RoboDK station: Robot_2_2025.rdk

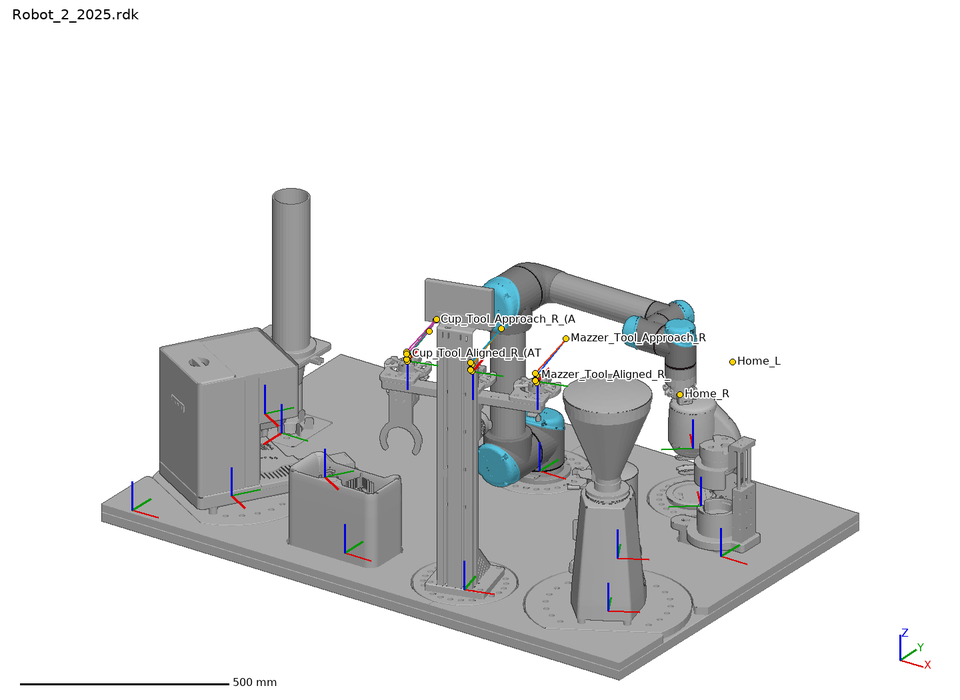
[picture v0: the station drawn from its stored meshes, robots at their saved joint values, targets as dots, program paths as lines]
Station Robot_2_2025 (saved by RoboDK 6.0.7). Poses are relative to the parent item; angles as X-Y-Z fixed-axis rotations.
Station parameters (name, value as stored): IO_5, 1, IO_2, 0, IO_3, 0, IO_4, 0, IO_1, 0, IO_0, 0, 0, 0, 1, 0, 4, 0
  - frame UR5_Base at (0, 0, 0) mm
    - robot UR5: 6 axes
        modified DH rows (alpha deg, a mm, theta deg, d mm): 0, 0, 0, 89.2; 90, 0, 180, 0; 0, 425, 0, 0; 0, 392, 0, 109.3; -90, 0, 0, 94.75; 90, 0, 180, 82.5
        joint limits [-360, -360, -360, -360, -360, -360] to [360, 360, 360, 360, 360, 360]; home [0, -90, -90, 0, 90, 0]; saved at [-0.001, -89.995, -89.998, -90.003, 89.998, 0.001]
      - tool Master_Tool_(UR5), TCP at (0, 0, 48.94) mm, size 88.9 x 94.7 x 67.9 mm
      - tool Cup_Tool_Shut_(UR5), TCP at (-34.39, 40.98, 235.56) mm, rotated rx 0 ry 0 rz -50 deg, size 116 x 104.2 x 218.8 mm
      - tool Cup_Tool_Open_(UR5), TCP at (-67.17, 80.05, 235.56) mm, rotated rx 0 ry 0 rz -50 deg, size 166.5 x 104.2 x 218.8 mm
      - tool Mazzer_Tool_(UR5), TCP at (0, 0, 153.18) mm, rotated rx 0 ry 0 rz -50 deg, size 105.5 x 104.2 x 106.6 mm
      - tool Rancilio_Tool_(UR5), TCP at (18.19, -21.68, 194.84) mm, rotated rx 0 ry -3.9 rz -50 deg, size 87.5 x 104.2 x 184.8 mm
      - tool Cup_(UR5), TCP at (-82.31, 98.09, 235.54) mm, rotated rx 0 ry 0 rz -50 deg, size 79 x 78 x 79 mm
    - object UR5_Plate at (0, 0, 0) mm, size 249.9 x 249.9 x 20 mm, geometry from UR5_Plate.STL
    - frame Table_Top at (-700, -700, -20) mm
      - object Table_Top at (0, 0, 0) mm, size 1515 x 1000 x 25 mm, geometry from Table_Top.STL
      - object Table_Cushion at (0, 0, 0) mm, size 1515 x 1000 x 20 mm, geometry from Table_Cushion.STL
      - frame Rancilio at (150, 200, 0) mm, rotated rx 0 ry 0 rz -30 deg
        - object Rancilio at (0, 0, 0) mm, size 399.6 x 458 x 388.3 mm, geometry from Rancilio_Assembly.STL
        - frame Rancilio_Tool at (39.29, 69.7, 222) mm
          - object Rancilio_Tool_Inserted_(Rancilio) at (0, 0, 0) mm, rotated rx 0 ry -90 rz 45 deg, size 87.1 x 104.3 x 184.1 mm, geometry from Rancilio_Tool_Assembly.STL
          - object Rancilio_Tool_Rotated_(Rancilio) at (0, 0, 0) mm, rotated rx 0 ry -90 rz 75 deg, size 87.1 x 104.3 x 184.1 mm, geometry from Rancilio_Tool_Assembly.STL
        - frame Rancilio_Scale at (39, 226.92, 20) mm
          - object Cup_(Rancilio) at (0, -157.52, 65.24) mm, size 79 x 79 x 78 mm, geometry from Supreme_Cup.STL
          - object Rancilio_Scale_Lock at (0, 0, 0) mm, size 100.1 x 260 x 71.4 mm, geometry from Rancilio_Scale_Assembly_1_Lock.STL
          - object Rancilio_Scale_Read at (0, 0, 0) mm, size 100.1 x 260 x 71.4 mm, geometry from Rancilio_Scale_Assembly_1_Read.STL
      - frame Rancilio_Tool_Cleaner at (550, 100, 0) mm
        - object Rancilio_Tool_Cleaner at (0, 0, 0) mm, size 258 x 136.9 x 218.7 mm, geometry from Portafilter_Cleaner_Assembly.STL
      - frame ATI at (900, 100, 0) mm, rotated rx 0 ry 0 rz 15 deg
        - object ATI at (0, 0, 0) mm, size 444.3 x 250 x 843.3 mm, geometry from ATI_Assembly_1.STL
        - frame Cup_Tool_(ATI) at (-163.9, 54.25, 556) mm, rotated rx 180 ry 0 rz 90 deg
          - object Cup_Tool_Shut_(ATI) at (0, 0, 0) mm, size 116 x 104.3 x 218.9 mm, geometry from Cup_Tool_Assembly_Closed.STL
          - target Cup_Tool_Approach_R_(ATI) (joint target) at (200, -1, -18) mm, rotated rx 0 ry 0 rz 50 deg; joints [-77.671, -81.541, -71.804, -116.654, 90.001, -222.671] of UR5
          - target Cup_Tool_Aligned_R_(ATI) (joint target) at (0.64, -1.17, -18.29) mm, rotated rx -0.48 ry 0.34 rz 50.01 deg; joints [-76.902, -110.177, -39.589, -120.099, 90.575, -221.892] of UR5
          - target Cup_Tool_Inserted_R_(ATI) (joint target) at (1.17, -1.09, 0) mm, rotated rx -0.52 ry 0.38 rz 50.08 deg; joints [-76.908, -108.351, -45.194, -116.323, 90.631, -221.828] of UR5
          - target Cup_Tool_Mated_R_(ATI) (joint target) at (0.72, -1.18, 0.85) mm, rotated rx -0.51 ry 0.38 rz 50.07 deg; joints [-76.914, -108.36, -45.32, -116.191, 90.623, -221.837] of UR5
          - target Cup_Tool_Attached_R_(ATI) (joint target) at (1.05, -1.02, -11) mm, rotated rx -0.5 ry 0.36 rz 50.03 deg; joints [-76.894, -109.363, -41.97, -118.536, 90.601, -221.86] of UR5
          - target Cup_Tool_Rotated_R_(ATI) (joint target) at (1.07, -1.03, -11.05) mm, rotated rx 0.35 ry 0.5 rz 140.04 deg; joints [-76.895, -109.361, -41.967, -118.536, 90.599, -131.856] of UR5
          - target Cup_Tool_Departure_R_(ATI) (joint target) at (151, -1, -11) mm, rotated rx 0 ry 0 rz 140 deg; joints [-77.368, -87.366, -67.792, -114.84, 90.001, -132.368] of UR5
          - target Cup_Tool_Approach_L_(ATI) (joint target) at (200, 0, -20) mm, rotated rx 0 ry 0 rz 50.44 deg; joints [70.564, -98.372, 71.405, -63.033, -89.998, -254] of UR5
          - target Cup_Tool_Aligned_L_(ATI) (joint target) at (2.26, -4.72, -23.42) mm, rotated rx -0.9 ry 0.14 rz 50.33 deg; joints [81.304, -69.621, 38.471, -59.135, -89.129, -243.367] of UR5
          - target Cup_Tool_Inserted_L_(ATI) (joint target) at (2, -4.79, -4.65) mm, rotated rx -0.97 ry 0.67 rz 50.05 deg; joints [81.242, -71.217, 43.754, -62.366, -88.837, -243.702] of UR5
          - target Cup_Tool_Mated_L_(ATI) (joint target) at (2.09, -4.82, -3.48) mm, rotated rx -0.94 ry 0.16 rz 50.41 deg; joints [81.293, -71.561, 44.547, -63.271, -89.089, -243.297] of UR5
          - target Cup_Tool_Attached_L_(ATI) (joint target) at (2.12, -4.74, -16.57) mm, rotated rx -0.94 ry 0.65 rz 50 deg; joints [81.249, -70.086, 40.174, -59.922, -88.864, -243.75] of UR5
          - target Cup_Tool_Rotated_L_(ATI) (joint target) at (2.13, -4.71, -16.62) mm, rotated rx 0.65 ry 0.95 rz 140.01 deg; joints [81.251, -70.088, 40.172, -59.924, -88.864, -153.749] of UR5
          - target Cup_Tool_Departure_L_(ATI) (joint target) at (151, -1, -11) mm, rotated rx 0 ry 0 rz 140 deg; joints [74.169, -92.634, 67.792, -65.159, -89.998, -160.831] of UR5
        - frame Mazzer_Tool_(ATI) at (165.9, 57.75, 555.5) mm, rotated rx 180 ry 0 rz 90 deg
          - object Mazzer_Tool_(ATI) at (0, 0, 0) mm, size 105.5 x 104.3 x 106.6 mm, geometry from Mazzer_Tool_Assembly.STL
          - target Mazzer_Tool_Approach_R_(ATI) (joint target) at (200, -1, -21.5) mm, rotated rx 0 ry 0 rz 50 deg; joints [-31.604, -85.352, -68.03, -116.616, 90, -176.604] of UR5
          - target Mazzer_Tool_Aligned_R_(ATI) (joint target) at (-4.5, -1, -18.5) mm, rotated rx 0 ry 0 rz 50 deg; joints [-45.391, -114.596, -33.046, -122.356, 90, -190.391] of UR5
          - target Mazzer_Tool_Inserted_R_(ATI) (joint target) at (-4.5, -1, -0.5) mm, rotated rx 0 ry 0 rz 50 deg; joints [-45.391, -112.519, -39.214, -118.265, 90, -190.391] of UR5
          - target Mazzer_Tool_Mated_R_(ATI) (joint target) at (-4.5, -1, 0.5) mm, rotated rx 0 ry 0 rz 50 deg; joints [-45.391, -112.419, -39.527, -118.052, 90, -190.391] of UR5
          - target Mazzer_Tool_Approach_L_(ATI) (joint target) at (200, -1, -21.5) mm, rotated rx 0 ry 0 rz 50 deg; joints [118.595, -94.648, 68.03, -63.384, -89.999, -206.405] of UR5
          - target Mazzer_Tool_Aligned_L_(ATI) (joint target) at (-4.36, -4.86, -23.14) mm, rotated rx -0.19 ry 0.13 rz 49.98 deg; joints [113.647, -65.161, 31.892, -56.831, -89.788, -211.369] of UR5
          - target Mazzer_Tool_Inserted_L_(ATI) (joint target) at (-4.52, -4.92, -5.11) mm, rotated rx -0.22 ry 0.17 rz 50.07 deg; joints [113.629, -67.327, 38.245, -61.015, -89.74, -211.299] of UR5
          - target Mazzer_Tool_Mated_L_(ATI) (joint target) at (-5.2, -5.01, -3.66) mm, rotated rx -0.41 ry 0.08 rz 50.34 deg; joints [113.605, -67.494, 38.794, -61.616, -89.718, -211.049] of UR5
        - frame Rancilio_Tool_(ATI) at (1, 56, 555.5) mm, rotated rx 180 ry 0 rz 90 deg
          - object Rancilio_Tool_(ATI) at (0, 0, 0) mm, size 87.5 x 104.3 x 184.8 mm, geometry from Rancilio_Tool_Assembly.STL
          - target Rancilio_Tool_Approach_R_(ATI) (joint target) at (200, -1, -21.5) mm, rotated rx 0 ry 0 rz 50 deg; joints [-52.392, -79.027, -73.308, -117.663, 90.001, -197.392] of UR5
          - target Rancilio_Tool_Aligned_R_(ATI) (joint target) at (-1.75, -1, -18.5) mm, rotated rx 0 ry 0 rz 50 deg; joints [-60.349, -108.011, -42.651, -119.336, 90.001, -205.349] of UR5
          - target Rancilio_Tool_Inserted_R_(ATI) (joint target) at (-1.75, -1, -0.5) mm, rotated rx 0 ry 0 rz 50 deg; joints [-60.349, -106.429, -47.774, -115.795, 90.001, -205.349] of UR5
          - target Rancilio_Tool_Mated_R_(ATI) (joint target) at (-1.75, -1, -0.9) mm, rotated rx 0 ry 0 rz 50 deg; joints [-60.349, -106.461, -47.667, -115.871, 90.001, -205.349] of UR5
          - target Rancilio_Tool_Approach_L_(ATI) (joint target) at (200, -1, -21.5) mm, rotated rx 0 ry 0 rz 50 deg; joints [93.922, -100.973, 73.308, -62.336, -89.999, -231.078] of UR5
          - target Rancilio_Tool_Aligned_L_(ATI) (joint target) at (-1.15, -4.84, -22.91) mm, rotated rx -0.46 ry -0.06 rz 50.35 deg; joints [97.401, -71.926, 41.922, -60.359, -89.702, -227.248] of UR5
          - target Rancilio_Tool_Inserted_L_(ATI) (joint target) at (-1.43, -4.76, -4.98) mm, rotated rx -0.29 ry 0.72 rz 50.05 deg; joints [97.32, -73.179, 46.429, -62.916, -89.302, -227.628] of UR5
          - target Rancilio_Tool_Mated_L_(ATI) (joint target) at (-1.31, -4.89, -4.19) mm, rotated rx -0.49 ry -0.04 rz 50.43 deg; joints [97.39, -73.597, 47.306, -64.072, -89.665, -227.181] of UR5
      - frame Mazzer at (1250, 200, 0) mm, rotated rx 0 ry 0 rz 30 deg
        - object Mazzer at (0, 0, 0) mm, size 399.9 x 495 x 614.6 mm, geometry from Mazzer_Assembly_1.STL
        - frame Mazzer_Scale at (0, 250, 20) mm
          - object Rancilio_Tool_(Mazzer) at (0, 40.18, 83.9) mm, rotated rx 0 ry -90 rz 90 deg, size 87.5 x 104.3 x 184.8 mm, geometry from Rancilio_Tool_Assembly.STL
          - object Mazzer_Scale_Lock at (0, 0, 0) mm, size 100.1 x 172.3 x 103.6 mm, geometry from Mazzer_Scale_Assembly_1_Lock.STL
          - object Mazzer_Scale_Read at (0, 0, 0) mm, size 100.1 x 172.3 x 103.6 mm, geometry from Mazzer_Scale_Assembly_1_Read.STL
      - frame Cup_Dispenser at (50, 550, 0) mm, rotated rx 0 ry 0 rz -90 deg
        - object Cup_Dispenser_Shut at (0, 0, 0) mm, size 162 x 208 x 656.6 mm, geometry from Cup_Dispenser_Assembly_Closed.STL
        - object Cup_Dispenser_Open at (0, 0, 0) mm, size 162 x 244.5 x 656.6 mm, geometry from Cup_Dispenser_Assembly_Open.STL
        - object Cup_(Cup_Dispenser) at (0, 27.5, 0) mm, size 79 x 79 x 78 mm, geometry from Supreme_Cup.STL
      - frame PUQ at (1100, 800, 0) mm, rotated rx 0 ry 0 rz 130 deg
        - object PUQ at (0, 0, 0) mm, size 249.7 x 250 x 301 mm, geometry from PUQ_Assembly.STL
        - frame Rancilio_Tool at (0, 18.5, 153.57) mm
          - object Rancilio_Tool_(PUQ) at (0, 0, 0) mm, rotated rx 0 ry -90 rz 90 deg, size 87.1 x 104.3 x 184.1 mm, geometry from Rancilio_Tool_Assembly.STL
      - frame WDT at (1300, 600, 0) mm
        - object Rancilio_Tool_(WDT) at (-10, 0, 133.57) mm, rotated rx 0 ry -90 rz -180 deg, size 87.1 x 104.3 x 184.1 mm, geometry from Rancilio_Tool_Assembly.STL
        - object WDT_Open at (0, 0, 0) mm, size 233 x 150 x 344.6 mm, geometry from UK_Tool_Assembly_Open.STL
        - object WDT_Shut at (0, 0, 0) mm, size 233 x 150 x 244.6 mm, geometry from UK_Tool_Assembly_Shut.STL
      - target Home_R (joint target) at (1186.72, 590.69, 402.81) mm, rotated rx -180 ry 0 rz -90 deg; joints [-0.001, -89.995, -89.998, -90.003, 89.998, 0.001] of UR5
      - target Home_L (joint target) at (1186.75, 809.3, 402.76) mm, rotated rx -180 ry 0 rz 0 deg; joints [180, -90, 90, -90, -90, -90] of UR5
  - folder Tool_Programs
    - program Cup_Tool_Attach_R_(ATI) (14 instructions, listed below)
    - program Cup_Tool_Attach_L_(ATI) (14 instructions, listed below)
    - program Cup_Tool_Detach_R_(ATI) (17 instructions, listed below)
    - program Cup_Tool_Detach_L_(ATI) (17 instructions, listed below)
    - program WDT_Open (6 instructions, listed below)
    - program WDT_Shut (6 instructions, listed below)
    - program Mazzer_Tool_Attach_R_(ATI) (12 instructions, listed below)
    - program Mazzer_Tool_Attach_L_(ATI) (12 instructions, listed below)
    - program Mazzer_Tool_Detach_R_(ATI) (16 instructions, listed below)
    - program Mazzer_Tool_Detach_L_(ATI) (16 instructions, listed below)
    - program Rancilio_Tool_Attach_R_(ATI) (12 instructions, listed below)
    - program Rancilio_Tool_Attach_L_(ATI) (12 instructions, listed below)
    - program Rancilio_Tool_Detach_R_(ATI) (15 instructions, listed below)
    - program Rancilio_Tool_Detach_L_(ATI) (15 instructions, listed below)
    - program Cup_Tool_Open_(UR5) (5 instructions, listed below)
    - program Cup_Tool_Shut_(UR5) (5 instructions, listed below)
    - program Student_Tool_Attach (2 instructions, listed below)
    - program Student_Tool_Detach (5 instructions, listed below)
  - folder Visual_Programs
    - program Reset_Simulation_L (25 instructions, listed below)
    - program Reset_Simulation_R (25 instructions, listed below)
    - program Show_Rancilio_Scale_Lock (2 instructions, listed below)
    - program Show_Rancilio_Scale_Read (2 instructions, listed below)
    - program Show_Mazzer_Scale_Lock (2 instructions, listed below)
    - program Show_Mazzer_Scale_Read (2 instructions, listed below)
    - program Show_Mazzer_Scale_Rancilio_Tool (1 instructions, listed below)
    - program Hide_Mazzer_Scale_Rancilio_Tool (1 instructions, listed below)
    - program Show_Rancilio_Scale_Cup (1 instructions, listed below)
    - program Hide_Rancilio_Scale_Cup (1 instructions, listed below)
    - program Show_Cup_Dispenser_Cup (1 instructions, listed below)
    - program Hide_Cup_Dispenser_Cup (1 instructions, listed below)
    - program Show_Cup_Dispenser_Open (2 instructions, listed below)
    - program Show_Cup_Dispenser_Shut (2 instructions, listed below)
    - program Show_WDT_Shut (2 instructions, listed below)
    - program Show_WDT_Open (2 instructions, listed below)
    - program Hide_WDT_Rancilio_Tool (1 instructions, listed below)
    - program Show_WDT_Rancilio_Tool (1 instructions, listed below)
    - program Show_Cup_Tool_Cup (1 instructions, listed below)
    - program Hide_Cup_Tool_Cup (1 instructions, listed below)
    - program Show_Rancilio_Rancilio_Tool_Rotated (1 instructions, listed below)
    - program Hide_Rancilio_Rancilio_Tool_Rotated (1 instructions, listed below)
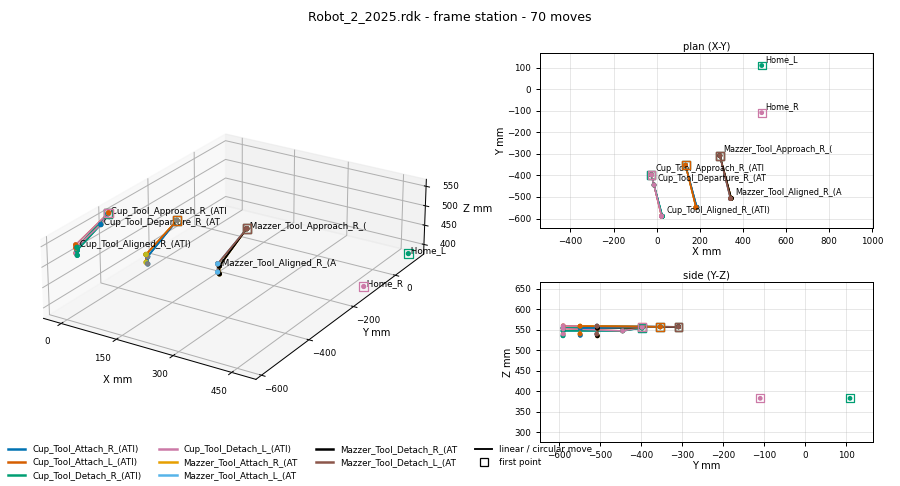
[picture p0: tool path of Robot_2_2025.rdk in frame station, 70 of 70 moves have a stored position in this frame; points joined in program order, loops and branches not executed]

--- program Cup_Tool_Attach_R_(ATI) (robot UR5) ---
  Set Ref.: Cup_Tool_(ATI)
  Set Tool: Master_Tool_(UR5)
  MoveJ (Cup_Tool_Approach_R_(ATI))
  MoveL (Cup_Tool_Aligned_R_(ATI))
  MoveL (Cup_Tool_Mated_R_(ATI))
  Set IO_0=1
  Pause 500 ms
  Hide Cup_Tool_Shut_(ATI)
  Show Cup_Tool_Shut_(UR5)
  MoveL (Cup_Tool_Attached_R_(ATI))
  MoveL (Cup_Tool_Rotated_R_(ATI))
  MoveL (Cup_Tool_Departure_R_(ATI))
  MoveL (Cup_Tool_Approach_R_(ATI))
  Set Ref.: UR5_Base

--- program Cup_Tool_Attach_L_(ATI) (robot UR5) ---
  Set Ref.: Cup_Tool_(ATI)
  Set Tool: Master_Tool_(UR5)
  MoveJ (Cup_Tool_Approach_L_(ATI))
  MoveL (Cup_Tool_Aligned_L_(ATI))
  MoveL (Cup_Tool_Mated_L_(ATI))
  Set IO_0=1
  Pause 500 ms
  Hide Cup_Tool_Shut_(ATI)
  Show Cup_Tool_Shut_(UR5)
  MoveL (Cup_Tool_Attached_L_(ATI))
  MoveL (Cup_Tool_Rotated_L_(ATI))
  MoveL (Cup_Tool_Departure_L_(ATI))
  MoveL (Cup_Tool_Approach_L_(ATI))
  Set Ref.: UR5_Base

--- program Cup_Tool_Detach_R_(ATI) (robot UR5) ---
  Set Ref.: Cup_Tool_(ATI)
  Set Tool: Master_Tool_(UR5)
  MoveJ (Cup_Tool_Approach_R_(ATI))
  MoveL (Cup_Tool_Departure_R_(ATI))
  MoveL (Cup_Tool_Rotated_R_(ATI))
  MoveL (Cup_Tool_Attached_R_(ATI))
  MoveL (Cup_Tool_Mated_R_(ATI))
  Set IO_0=0
  Pause 500 ms
  Set IO_1=1
  Pause 500 ms
  Set IO_1=0
  Hide Cup_Tool_Shut_(UR5)
  Show Cup_Tool_Shut_(ATI)
  MoveL (Cup_Tool_Aligned_R_(ATI))
  MoveL (Cup_Tool_Approach_R_(ATI))
  Set Ref.: UR5_Base

--- program Cup_Tool_Detach_L_(ATI) (robot UR5) ---
  Set Ref.: Cup_Tool_(ATI)
  Set Tool: Master_Tool_(UR5)
  MoveJ (Cup_Tool_Approach_L_(ATI))
  MoveL (Cup_Tool_Departure_L_(ATI))
  MoveL (Cup_Tool_Rotated_L_(ATI))
  MoveL (Cup_Tool_Attached_L_(ATI))
  MoveL (Cup_Tool_Mated_L_(ATI))
  Set IO_0=0
  Pause 500 ms
  Set IO_1=1
  Pause 500 ms
  Set IO_1=0
  Hide Cup_Tool_Shut_(UR5)
  Show Cup_Tool_Shut_(ATI)
  MoveL (Cup_Tool_Aligned_L_(ATI))
  MoveL (Cup_Tool_Approach_L_(ATI))
  Set Ref.: UR5_Base

--- program WDT_Open (robot UR5) ---
  Set IO_4=1
  Pause 500 ms
  Set IO_4=0
  Pause 500 ms
  Hide WDT_Shut
  Show WDT_Open

--- program WDT_Shut (robot UR5) ---
  Set IO_5=1
  Pause 500 ms
  Set IO_5=0
  Pause 500 ms
  Hide WDT_Open
  Show WDT_Shut

--- program Mazzer_Tool_Attach_R_(ATI) (robot UR5) ---
  Set Ref.: Mazzer_Tool_(ATI)
  Set Tool: Master_Tool_(UR5)
  MoveJ (Mazzer_Tool_Approach_R_(ATI))
  MoveL (Mazzer_Tool_Aligned_R_(ATI))
  MoveL (Mazzer_Tool_Mated_R_(ATI))
  Set IO_0=1
  Pause 500 ms
  Hide Mazzer_Tool_(ATI)
  Show Mazzer_Tool_(UR5)
  MoveL (Mazzer_Tool_Aligned_R_(ATI))
  MoveL (Mazzer_Tool_Approach_R_(ATI))
  Set Ref.: UR5_Base

--- program Mazzer_Tool_Attach_L_(ATI) (robot UR5) ---
  Set Ref.: Mazzer_Tool_(ATI)
  Set Tool: Master_Tool_(UR5)
  MoveJ (Mazzer_Tool_Approach_L_(ATI))
  MoveL (Mazzer_Tool_Aligned_L_(ATI))
  MoveL (Mazzer_Tool_Mated_L_(ATI))
  Set IO_0=1
  Pause 500 ms
  Hide Mazzer_Tool_(ATI)
  Show Mazzer_Tool_(UR5)
  MoveL (Mazzer_Tool_Aligned_L_(ATI))
  MoveL (Mazzer_Tool_Approach_L_(ATI))
  Set Ref.: UR5_Base

--- program Mazzer_Tool_Detach_R_(ATI) (robot UR5) ---
  Set Ref.: Mazzer_Tool_(ATI)
  Set Tool: Master_Tool_(UR5)
  MoveJ (Mazzer_Tool_Approach_R_(ATI))
  MoveL (Mazzer_Tool_Aligned_R_(ATI))
  MoveL (Mazzer_Tool_Mated_R_(ATI))
  Set IO_0=0
  Pause 500 ms
  Set IO_1=1
  Pause 500 ms
  Set IO_1=0
  Hide Mazzer_Tool_(UR5)
  Show Mazzer_Tool_(ATI)
  MoveL (Mazzer_Tool_Aligned_R_(ATI))
  MoveL (Mazzer_Tool_Approach_R_(ATI))
  Set Ref.: UR5_Base
  Set Tool: Master_Tool_(UR5)

--- program Mazzer_Tool_Detach_L_(ATI) (robot UR5) ---
  Set Ref.: Mazzer_Tool_(ATI)
  Set Tool: Master_Tool_(UR5)
  MoveJ (Mazzer_Tool_Approach_L_(ATI))
  MoveL (Mazzer_Tool_Aligned_L_(ATI))
  MoveL (Mazzer_Tool_Mated_L_(ATI))
  Set IO_0=0
  Pause 500 ms
  Set IO_1=1
  Pause 500 ms
  Set IO_1=0
  Hide Mazzer_Tool_(UR5)
  Show Mazzer_Tool_(ATI)
  MoveL (Mazzer_Tool_Aligned_L_(ATI))
  MoveL (Mazzer_Tool_Approach_L_(ATI))
  Set Ref.: UR5_Base
  Set Tool: Master_Tool_(UR5)

--- program Rancilio_Tool_Attach_R_(ATI) (robot UR5) ---
  Set Ref.: Rancilio_Tool_(ATI)
  Set Tool: Master_Tool_(UR5)
  MoveJ (Rancilio_Tool_Approach_R_(ATI))
  MoveL (Rancilio_Tool_Aligned_R_(ATI))
  MoveL (Rancilio_Tool_Mated_R_(ATI))
  Set IO_0=1
  Pause 500 ms
  Hide Rancilio_Tool_(ATI)
  Show Rancilio_Tool_(UR5)
  MoveL (Rancilio_Tool_Aligned_R_(ATI))
  MoveL (Rancilio_Tool_Approach_R_(ATI))
  Set Ref.: UR5_Base

--- program Rancilio_Tool_Attach_L_(ATI) (robot UR5) ---
  Set Ref.: Rancilio_Tool_(ATI)
  Set Tool: Master_Tool_(UR5)
  MoveJ (Rancilio_Tool_Approach_L_(ATI))
  MoveL (Rancilio_Tool_Aligned_L_(ATI))
  MoveL (Rancilio_Tool_Mated_L_(ATI))
  Set IO_0=1
  Pause 500 ms
  Hide Rancilio_Tool_(ATI)
  Show Rancilio_Tool_(UR5)
  MoveL (Rancilio_Tool_Aligned_L_(ATI))
  MoveL (Rancilio_Tool_Approach_L_(ATI))
  Set Ref.: UR5_Base

--- program Rancilio_Tool_Detach_R_(ATI) (robot UR5) ---
  Set Ref.: Rancilio_Tool_(ATI)
  Set Tool: Master_Tool_(UR5)
  MoveJ (Rancilio_Tool_Approach_R_(ATI))
  MoveL (Rancilio_Tool_Aligned_R_(ATI))
  MoveL (Rancilio_Tool_Mated_R_(ATI))
  Set IO_0=0
  Pause 500 ms
  Set IO_1=1
  Pause 500 ms
  Set IO_1=0
  Hide Rancilio_Tool_(UR5)
  Show Rancilio_Tool_(ATI)
  MoveL (Rancilio_Tool_Aligned_R_(ATI))
  MoveL (Rancilio_Tool_Approach_R_(ATI))
  Set Ref.: UR5_Base

--- program Rancilio_Tool_Detach_L_(ATI) (robot UR5) ---
  Set Ref.: Rancilio_Tool_(ATI)
  Set Tool: Master_Tool_(UR5)
  MoveJ (Rancilio_Tool_Approach_L_(ATI))
  MoveL (Rancilio_Tool_Aligned_L_(ATI))
  MoveL (Rancilio_Tool_Mated_L_(ATI))
  Set IO_0=0
  Pause 500 ms
  Set IO_1=1
  Pause 500 ms
  Set IO_1=0
  Hide Rancilio_Tool_(UR5)
  Show Rancilio_Tool_(ATI)
  MoveL (Rancilio_Tool_Aligned_L_(ATI))
  MoveL (Rancilio_Tool_Approach_L_(ATI))
  Set Ref.: UR5_Base

--- program Cup_Tool_Open_(UR5) (robot UR5) ---
  Set IO_2=1
  Hide Cup_Tool_Shut_(UR5)
  Show Cup_Tool_Open_(UR5)
  Pause 500 ms
  Set IO_2=0

--- program Cup_Tool_Shut_(UR5) (robot UR5) ---
  Set IO_3=1
  Hide Cup_Tool_Open_(UR5)
  Show Cup_Tool_Shut_(UR5)
  Pause 500 ms
  Set IO_3=0

--- program Student_Tool_Attach (robot UR5) ---
  Set IO_0=1
  Pause 500 ms

--- program Student_Tool_Detach (robot UR5) ---
  Set IO_0=0
  Pause 500 ms
  Set IO_1=1
  Pause 500 ms
  Set IO_1=0

--- program Reset_Simulation_L (robot UR5) ---
  MoveJ (Home_L)
  Show Master_Tool_(UR5)
  Hide Cup_Tool_Shut_(UR5)
  Hide Cup_Tool_Open_(UR5)
  Hide Mazzer_Tool_(UR5)
  Hide Rancilio_Tool_(UR5)
  Hide Cup_(UR5)
  Hide Rancilio_Tool_Inserted_(Rancilio)
  Hide Rancilio_Tool_Rotated_(Rancilio)
  Hide Cup_(Rancilio)
  Hide Rancilio_Scale_Read
  Show Rancilio_Scale_Lock
  Show Cup_Tool_Shut_(ATI)
  Show Mazzer_Tool_(ATI)
  Show Rancilio_Tool_(ATI)
  Hide Mazzer_Scale_Read
  Show Mazzer_Scale_Lock
  Hide Cup_Dispenser_Open
  Show Cup_Dispenser_Shut
  Hide Cup_(Cup_Dispenser)
  Hide Rancilio_Tool_(PUQ)
  Hide Rancilio_Tool_(Mazzer)
  Hide WDT_Open
  Show WDT_Shut
  Hide Rancilio_Tool_(WDT)

--- program Reset_Simulation_R (robot UR5) ---
  MoveJ (Home_R)
  Show Master_Tool_(UR5)
  Hide Cup_Tool_Shut_(UR5)
  Hide Cup_Tool_Open_(UR5)
  Hide Mazzer_Tool_(UR5)
  Hide Rancilio_Tool_(UR5)
  Hide Cup_(UR5)
  Hide Rancilio_Tool_Inserted_(Rancilio)
  Hide Rancilio_Tool_Rotated_(Rancilio)
  Hide Cup_(Rancilio)
  Hide Rancilio_Scale_Read
  Show Rancilio_Scale_Lock
  Show Cup_Tool_Shut_(ATI)
  Show Mazzer_Tool_(ATI)
  Show Rancilio_Tool_(ATI)
  Hide Mazzer_Scale_Read
  Show Mazzer_Scale_Lock
  Hide Cup_Dispenser_Open
  Show Cup_Dispenser_Shut
  Hide Cup_(Cup_Dispenser)
  Hide Rancilio_Tool_(PUQ)
  Hide Rancilio_Tool_(Mazzer)
  Hide WDT_Open
  Show WDT_Shut
  Hide Rancilio_Tool_(WDT)

--- program Show_Rancilio_Scale_Lock (robot UR5) ---
  Show Rancilio_Scale_Lock
  Hide Rancilio_Scale_Read

--- program Show_Rancilio_Scale_Read (robot UR5) ---
  Hide Rancilio_Scale_Lock
  Show Rancilio_Scale_Read

--- program Show_Mazzer_Scale_Lock (robot UR5) ---
  Hide Mazzer_Scale_Read
  Show Mazzer_Scale_Lock

--- program Show_Mazzer_Scale_Read (robot UR5) ---
  Hide Mazzer_Scale_Lock
  Show Mazzer_Scale_Read

--- program Show_Mazzer_Scale_Rancilio_Tool (robot UR5) ---
  Show Rancilio_Tool_(Mazzer)

--- program Hide_Mazzer_Scale_Rancilio_Tool (robot UR5) ---
  Hide Rancilio_Tool_(Mazzer)

--- program Show_Rancilio_Scale_Cup (robot UR5) ---
  Show Cup_(Rancilio)

--- program Hide_Rancilio_Scale_Cup (robot UR5) ---
  Hide Cup_(Rancilio)

--- program Show_Cup_Dispenser_Cup (robot UR5) ---
  Show Cup_(Cup_Dispenser)

--- program Hide_Cup_Dispenser_Cup (robot UR5) ---
  Hide Cup_(Cup_Dispenser)

--- program Show_Cup_Dispenser_Open (robot UR5) ---
  Hide Cup_Dispenser_Shut
  Show Cup_Dispenser_Open

--- program Show_Cup_Dispenser_Shut (robot UR5) ---
  Hide Cup_Dispenser_Open
  Show Cup_Dispenser_Shut

--- program Show_WDT_Shut (robot UR5) ---
  Hide WDT_Open
  Show WDT_Shut

--- program Show_WDT_Open (robot UR5) ---
  Hide WDT_Shut
  Show WDT_Open

--- program Hide_WDT_Rancilio_Tool (robot UR5) ---
  Hide Rancilio_Tool_(WDT)

--- program Show_WDT_Rancilio_Tool (robot UR5) ---
  Show Rancilio_Tool_(WDT)

--- program Show_Cup_Tool_Cup (robot UR5) ---
  Show Cup_(UR5)

--- program Hide_Cup_Tool_Cup (robot UR5) ---
  Hide Cup_(UR5)

--- program Show_Rancilio_Rancilio_Tool_Rotated (robot UR5) ---
  Show Rancilio_Tool_Rotated_(Rancilio)

--- program Hide_Rancilio_Rancilio_Tool_Rotated (robot UR5) ---
  Hide Rancilio_Tool_Rotated_(Rancilio)
